TYPE "FRK_HealthBook"
VERSION : 0.1
   STRUCT
      "Slots" {ExternalAccessible := 'False'; ExternalVisible := 'False'; ExternalWritable := 'False'} : Array[1..12] of Int;
   END_STRUCT;
END_TYPE
